TYPE stSwitchState :
STRUCT
    StateType : eSwitchStateType;         // Current processed state
    PressCount : USINT := 0;            // Number of clicks in sequence
END_STRUCT
END_TYPE

(* stored: Version 1.1.0.1
   DUT stSwitchState: Id {95f89ab6-dc0c-4e63-95ce-633bc21eb204} *)
